// TIA Portal V20 export
FUNCTION_BLOCK "FB_LD_PressDemoHome"   // FB, LAD
{ S7_Optimized_Access := 'TRUE' }
// stored: AutoNumber true
   VAR_INPUT
      Run { ExternalWritable := 'False'} : Bool;
      Reset { ExternalWritable := 'False'} : Bool;
      OwnerIndex { ExternalWritable := 'False'} : DInt;
      Delta { ExternalWritable := 'False'} : Time;
   END_VAR
   VAR_IN_OUT
      PressRam { ExternalAccessible := 'False'; ExternalVisible := 'False'; ExternalWritable := 'False'} : "FB_CylinderCM";
      Door { ExternalAccessible := 'False'; ExternalVisible := 'False'; ExternalWritable := 'False'} : "FB_CylinderCM";
      PartSlide { ExternalAccessible := 'False'; ExternalVisible := 'False'; ExternalWritable := 'False'} : "FB_CylinderCM";
   END_VAR
   VAR
      Seq { ExternalWritable := 'False'} : "FRK_SequenceCtx";
      Row1 { ExternalWritable := 'False'} : "FRK_SequenceRow";
      Row2 { ExternalWritable := 'False'} : "FRK_SequenceRow";
      Row3 { ExternalWritable := 'False'} : "FRK_SequenceRow";
      Row4 { ExternalWritable := 'False'} : "FRK_SequenceRow";
      At0 { ExternalAccessible := 'False'; ExternalVisible := 'False'; ExternalWritable := 'False'} : Bool;
      At900 { ExternalAccessible := 'False'; ExternalVisible := 'False'; ExternalWritable := 'False'} : Bool;
      At910 { ExternalAccessible := 'False'; ExternalVisible := 'False'; ExternalWritable := 'False'} : Bool;
      At999 { ExternalAccessible := 'False'; ExternalVisible := 'False'; ExternalWritable := 'False'} : Bool;
      Ready1 { ExternalAccessible := 'False'; ExternalVisible := 'False'; ExternalWritable := 'False'} : Bool;
      Ready2 { ExternalAccessible := 'False'; ExternalVisible := 'False'; ExternalWritable := 'False'} : Bool;
      Ready3 { ExternalAccessible := 'False'; ExternalVisible := 'False'; ExternalWritable := 'False'} : Bool;
      Ready4 { ExternalAccessible := 'False'; ExternalVisible := 'False'; ExternalWritable := 'False'} : Bool;
      Ready5 { ExternalAccessible := 'False'; ExternalVisible := 'False'; ExternalWritable := 'False'} : Bool;
      Advance { ExternalAccessible := 'False'; ExternalVisible := 'False'; ExternalWritable := 'False'} : Bool;
   END_VAR
BEGIN

REGION Network 1
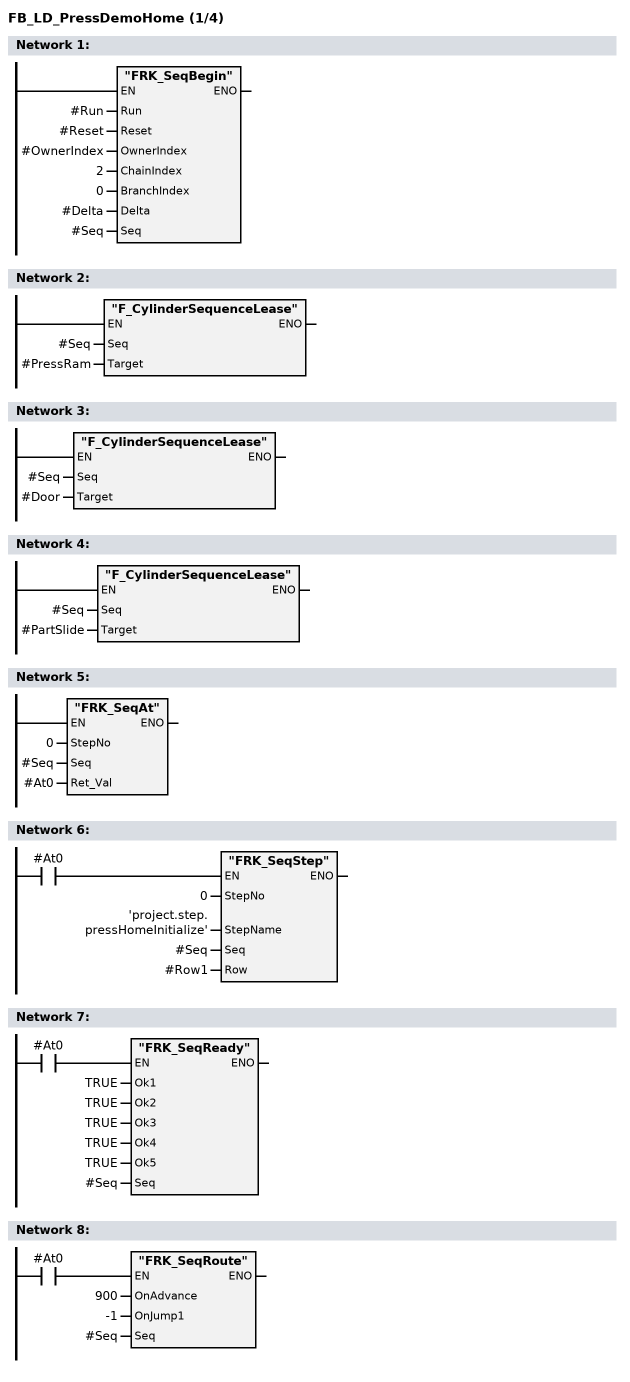
   RUNG wire#powerrail
      "FRK_SeqBegin"(Run := #Run, Reset := #Reset, OwnerIndex := #OwnerIndex, ChainIndex := 2, BranchIndex := 0, Delta := #Delta, Seq := #Seq)
   END_RUNG
   // the same network as SCL:
   "FRK_SeqBegin"(Run := #Run,
                  Reset := #Reset,
                  OwnerIndex := #OwnerIndex,
                  ChainIndex := 2,
                  BranchIndex := 0,
                  Delta := #Delta,
                  Seq := #Seq);
END_REGION

REGION Network 2
   RUNG wire#powerrail
      "F_CylinderSequenceLease"(Seq := #Seq, Target := #PressRam)
   END_RUNG
   // the same network as SCL:
   "F_CylinderSequenceLease"(Seq := #Seq, Target := #PressRam);
END_REGION

REGION Network 3
   RUNG wire#powerrail
      "F_CylinderSequenceLease"(Seq := #Seq, Target := #Door)
   END_RUNG
   // the same network as SCL:
   "F_CylinderSequenceLease"(Seq := #Seq, Target := #Door);
END_REGION

REGION Network 4
   RUNG wire#powerrail
      "F_CylinderSequenceLease"(Seq := #Seq, Target := #PartSlide)
   END_RUNG
   // the same network as SCL:
   "F_CylinderSequenceLease"(Seq := #Seq, Target := #PartSlide);
END_REGION

REGION Network 5
   RUNG wire#powerrail
      "FRK_SeqAt"(StepNo := 0, Seq := #Seq, Ret_Val := #At0)
   END_RUNG
   // the same network as SCL:
   "FRK_SeqAt"(StepNo := 0, Seq := #Seq, Ret_Val := #At0);
END_REGION

REGION Network 6
   IF #At0 THEN
       "FRK_SeqStep"(StepNo := 0, StepName := 'project.step.pressHomeInitialize', Seq := #Seq, Row := #Row1);
   END_IF;
END_REGION

REGION Network 7
   IF #At0 THEN
       "FRK_SeqReady"(Ok1 := TRUE, Ok2 := TRUE, Ok3 := TRUE, Ok4 := TRUE, Ok5 := TRUE, Seq := #Seq);
   END_IF;
END_REGION

REGION Network 8
   IF #At0 THEN "FRK_SeqRoute"(OnAdvance := 900, OnJump1 := -1, Seq := #Seq); END_IF;
END_REGION

REGION Network 9
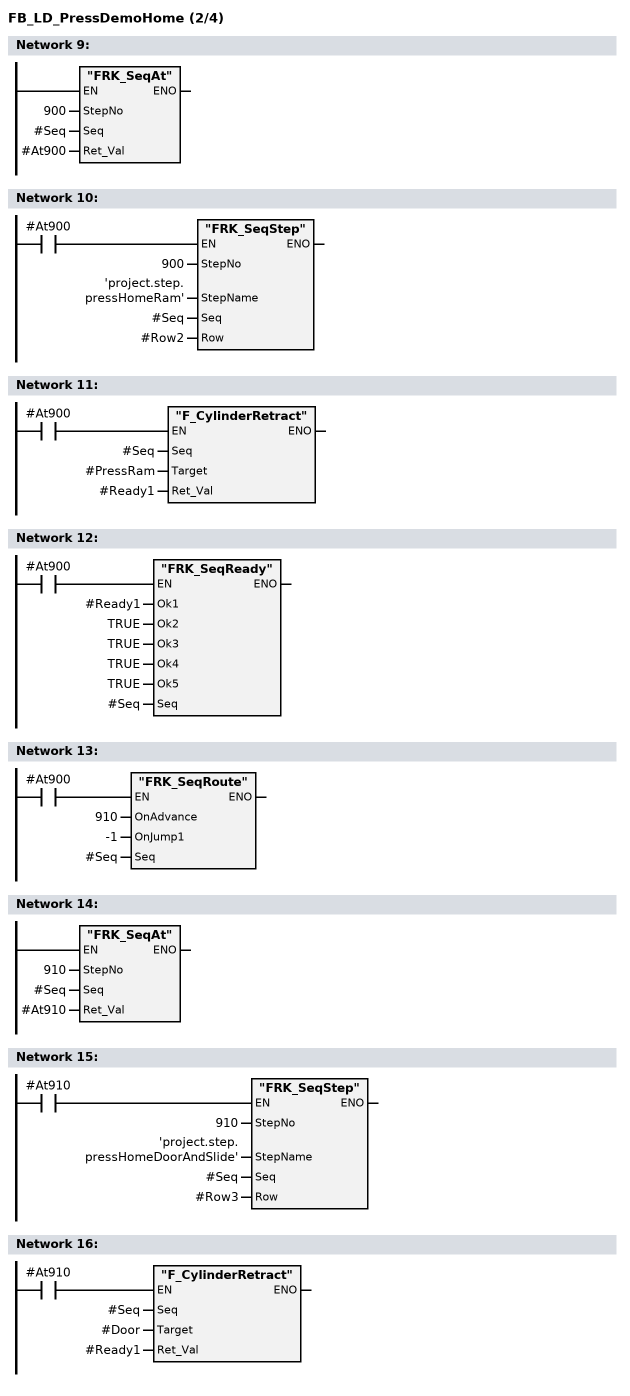
   RUNG wire#powerrail
      "FRK_SeqAt"(StepNo := 900, Seq := #Seq, Ret_Val := #At900)
   END_RUNG
   // the same network as SCL:
   "FRK_SeqAt"(StepNo := 900, Seq := #Seq, Ret_Val := #At900);
END_REGION

REGION Network 10
   IF #At900 THEN
       "FRK_SeqStep"(StepNo := 900, StepName := 'project.step.pressHomeRam', Seq := #Seq, Row := #Row2);
   END_IF;
END_REGION

REGION Network 11
   IF #At900 THEN "F_CylinderRetract"(Seq := #Seq, Target := #PressRam, Ret_Val := #Ready1); END_IF;
END_REGION

REGION Network 12
   IF #At900 THEN
       "FRK_SeqReady"(Ok1 := #Ready1, Ok2 := TRUE, Ok3 := TRUE, Ok4 := TRUE, Ok5 := TRUE, Seq := #Seq);
   END_IF;
END_REGION

REGION Network 13
   IF #At900 THEN "FRK_SeqRoute"(OnAdvance := 910, OnJump1 := -1, Seq := #Seq); END_IF;
END_REGION

REGION Network 14
   RUNG wire#powerrail
      "FRK_SeqAt"(StepNo := 910, Seq := #Seq, Ret_Val := #At910)
   END_RUNG
   // the same network as SCL:
   "FRK_SeqAt"(StepNo := 910, Seq := #Seq, Ret_Val := #At910);
END_REGION

REGION Network 15
   IF #At910 THEN
       "FRK_SeqStep"(StepNo := 910, StepName := 'project.step.pressHomeDoorAndSlide', Seq := #Seq, Row := #Row3);
   END_IF;
END_REGION

REGION Network 16
   IF #At910 THEN "F_CylinderRetract"(Seq := #Seq, Target := #Door, Ret_Val := #Ready1); END_IF;
END_REGION

REGION Network 17
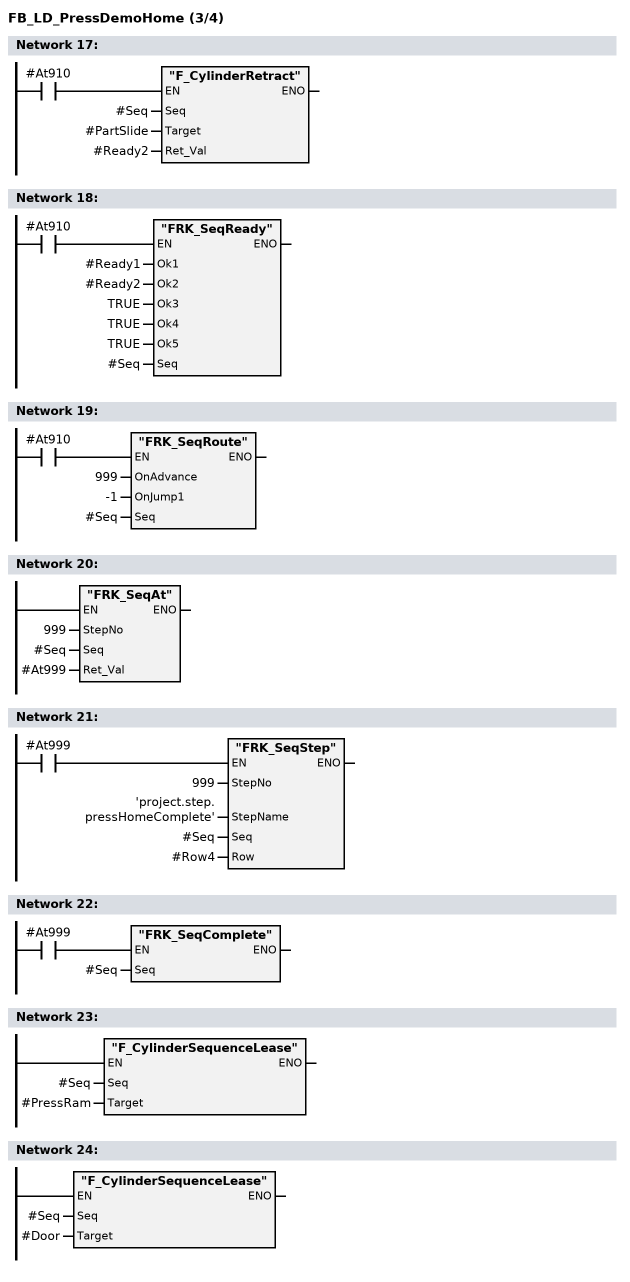
   IF #At910 THEN "F_CylinderRetract"(Seq := #Seq, Target := #PartSlide, Ret_Val := #Ready2); END_IF;
END_REGION

REGION Network 18
   IF #At910 THEN
       "FRK_SeqReady"(Ok1 := #Ready1, Ok2 := #Ready2, Ok3 := TRUE, Ok4 := TRUE, Ok5 := TRUE, Seq := #Seq);
   END_IF;
END_REGION

REGION Network 19
   IF #At910 THEN "FRK_SeqRoute"(OnAdvance := 999, OnJump1 := -1, Seq := #Seq); END_IF;
END_REGION

REGION Network 20
   RUNG wire#powerrail
      "FRK_SeqAt"(StepNo := 999, Seq := #Seq, Ret_Val := #At999)
   END_RUNG
   // the same network as SCL:
   "FRK_SeqAt"(StepNo := 999, Seq := #Seq, Ret_Val := #At999);
END_REGION

REGION Network 21
   IF #At999 THEN
       "FRK_SeqStep"(StepNo := 999, StepName := 'project.step.pressHomeComplete', Seq := #Seq, Row := #Row4);
   END_IF;
END_REGION

REGION Network 22
   IF #At999 THEN "FRK_SeqComplete"(Seq := #Seq); END_IF;
END_REGION

REGION Network 23
   RUNG wire#powerrail
      "F_CylinderSequenceLease"(Seq := #Seq, Target := #PressRam)
   END_RUNG
   // the same network as SCL:
   "F_CylinderSequenceLease"(Seq := #Seq, Target := #PressRam);
END_REGION

REGION Network 24
   RUNG wire#powerrail
      "F_CylinderSequenceLease"(Seq := #Seq, Target := #Door)
   END_RUNG
   // the same network as SCL:
   "F_CylinderSequenceLease"(Seq := #Seq, Target := #Door);
END_REGION

REGION Network 25
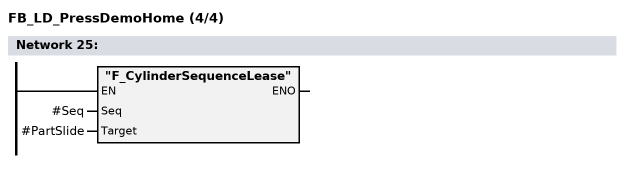
   RUNG wire#powerrail
      "F_CylinderSequenceLease"(Seq := #Seq, Target := #PartSlide)
   END_RUNG
   // the same network as SCL:
   "F_CylinderSequenceLease"(Seq := #Seq, Target := #PartSlide);
END_REGION
END_FUNCTION_BLOCK
